(* IEC 61131-3 sources: llm-plc-st-eval/data/processed/claude-sonnet-4-6/I6/zero_shot, 3 files *)

(* ---- ejec_3.st ---- *)
FUNCTION_BLOCK FB_Temperatura
VAR_INPUT
    rawTemp : INT;  (* Valor crudo del sensor: 0..27648 -> 0.0..100.0 °C *)
END_VAR

VAR_OUTPUT
    tempC     : REAL;  (* Temperatura calculada en grados Celsius *)
    enfriador : BOOL;  (* TRUE = enfriador activo *)
    almSensor : BOOL;  (* TRUE = señal fuera de rango *)
END_VAR

VAR CONSTANT
    RAW_MIN   : INT  := 0;       (* Valor crudo mínimo *)
    RAW_MAX   : INT  := 27648;   (* Valor crudo máximo *)
    TEMP_MIN  : REAL := 0.0;     (* Temperatura mínima en °C *)
    TEMP_MAX  : REAL := 100.0;   (* Temperatura máxima en °C *)
    HYST_HIGH : REAL := 80.0;    (* Umbral superior: activa enfriador *)
    HYST_LOW  : REAL := 75.0;    (* Umbral inferior: desactiva enfriador *)
END_VAR

(* ------------------------------------------------------------------ *)
(* 1. Verificación de rango del sensor                                 *)
(* ------------------------------------------------------------------ *)
IF rawTemp < RAW_MIN OR rawTemp > RAW_MAX THEN
    almSensor := TRUE;   (* Señal fuera de rango: alarma activa *)
    enfriador := FALSE;  (* Apagar enfriador por seguridad *)
    (* tempC conserva el último valor válido calculado *)
    RETURN;              (* Salir sin procesar más lógica *)
END_IF;

(* Sin alarma de sensor *)
almSensor := FALSE;

(* ------------------------------------------------------------------ *)
(* 2. Escalado lineal: rawTemp -> tempC                                *)
(*    tempC = (rawTemp - RAW_MIN) / (RAW_MAX - RAW_MIN) * TEMP_MAX    *)
(* ------------------------------------------------------------------ *)
tempC := (INT_TO_REAL(rawTemp) - INT_TO_REAL(RAW_MIN))
         / (INT_TO_REAL(RAW_MAX) - INT_TO_REAL(RAW_MIN))
         * (TEMP_MAX - TEMP_MIN)
         + TEMP_MIN;

(* ------------------------------------------------------------------ *)
(* 3. Control con histéresis del enfriador                             *)
(*    >= 80.0 °C -> encender  |  <= 75.0 °C -> apagar                 *)
(*    Entre 75.0 y 80.0 °C   -> mantener estado anterior              *)
(* ------------------------------------------------------------------ *)
IF tempC >= HYST_HIGH THEN
    enfriador := TRUE;   (* Temperatura alta: activar enfriador *)
ELSIF tempC <= HYST_LOW THEN
    enfriador := FALSE;  (* Temperatura baja: desactivar enfriador *)
(* ELSE: zona de histéresis, enfriador conserva su estado *)
END_IF;

(* ---- ejec_1.st ---- *)
(* ── Cuerpo del FUNCTION_BLOCK ── *)

(* 1. Verificar rango válido del sensor *)
IF rawTemp < RAW_MIN OR rawTemp > RAW_MAX THEN

    almSensor := TRUE;   (* Activar alarma de sensor fuera de rango *)
    enfriador := FALSE;  (* Desactivar enfriador por seguridad *)
    tempC     := 0.0;    (* Valor de temperatura indefinido, se fuerza a 0 *)

ELSE

    (* 2. Sin alarma: señal dentro de rango *)
    almSensor := FALSE;

    (* 3. Escalar rawTemp a grados Celsius (regla de tres lineal)
          tempC = (rawTemp - RAW_MIN) / (RAW_MAX - RAW_MIN) * (TEMP_MAX - TEMP_MIN) + TEMP_MIN
          Simplificado: tempC = rawTemp * 100.0 / 27648.0                              *)
    tempC := REAL_TO_REAL(INT_TO_REAL(rawTemp)) * (TEMP_MAX - TEMP_MIN)
             / INT_TO_REAL(RAW_MAX - RAW_MIN) + TEMP_MIN;

    (* 4. Control con histéresis (biestable):
          - Activa enfriador si tempC >= HYST_HIGH
          - Desactiva enfriador si tempC <= HYST_LOW
          - Entre ambos umbrales conserva el estado anterior (sin oscilar) *)
    IF tempC >= HYST_HIGH THEN
        enfriador := TRUE;
    ELSIF tempC <= HYST_LOW THEN
        enfriador := FALSE;
    (* ELSE: zona de histéresis -> enfriador mantiene su estado previo *)
    END_IF;

END_IF;

(* ---- ejec_2.st ---- *)
(* ── Cuerpo del bloque ─────────────────────────────────────────────────── *)

(* 1. Verificar rango del sensor *)
IF rawTemp < RAW_MIN OR rawTemp > RAW_MAX THEN

    almSensor := TRUE;   (* Activar alarma de sensor *)
    enfriador := FALSE;  (* Apagar enfriador por seguridad *)
    tempC     := 0.0;    (* Valor de temperatura indefinido → forzar a 0 *)

ELSE

    (* 2. Sin alarma de sensor *)
    almSensor := FALSE;

    (* 3. Escalar valor crudo a temperatura:
          tempC = (rawTemp - RAW_MIN) / (RAW_MAX - RAW_MIN) * (TEMP_MAX - TEMP_MIN) + TEMP_MIN
          Con RAW_MIN = 0 y TEMP_MIN = 0 se simplifica a:
          tempC = rawTemp / 27648.0 * 100.0                                *)
    tempC := (REAL#1.0 * rawTemp / REAL#27648.0) * (TEMP_MAX - TEMP_MIN) + TEMP_MIN;

    (* 4. Control con histéresis:
          - Activar  enfriador si tempC >= HYST_ON  (80.0 °C)
          - Desactivar         si tempC <= HYST_OFF (75.0 °C)
          - Entre ambos umbrales: conservar estado anterior (sin cambio)   *)
    IF tempC >= HYST_ON THEN
        enfriador := TRUE;
    ELSIF tempC <= HYST_OFF THEN
        enfriador := FALSE;
    (* ELSE: zona de histéresis → enfriador mantiene su estado actual *)
    END_IF;

END_IF;
